Fanuc KAREL source: KB00012.KL

PROGRAM KB00012
%NOLOCKGROUP
%ENVIRONMENT TPE
VAR
  P1: INTEGER
  P2: INTEGER
  P3: INTEGER
BEGIN
  P1 = 1
  P2 = 1
  P3 = 1
  AVL_POS_NUM(P1, P2, P3)
END KB00012
